(* IEC 61131-3 sources: plc-vscode/tests/st/test-ready/trust-platform/examples/OSCAT/tank_level_pid/non-oop/src, 3 files *)

(* ---- Configuration.st ---- *)
CONFIGURATION TankLevelPidClassicConfiguration
RESOURCE Cpu0 ON PLC
    TASK MainTask (INTERVAL := T#100ms, PRIORITY := 1);
    PROGRAM Main WITH MainTask : Main;
END_RESOURCE
END_CONFIGURATION

(* ---- Main.st ---- *)
PROGRAM Main
VAR
    TankController : CTRL_PID;
    LevelPercent : REAL := REAL#42.0;
    TargetLevelPercent : REAL := REAL#75.0;
    ValveCommandPercent : REAL;
    CommandLimited : BOOL;
END_VAR

TankController(
    ACT := LevelPercent,
    SET_POINT := TargetLevelPercent,
    SUP := REAL#0.0,
    OFS := REAL#0.0,
    M_I := REAL#35.0,
    MAN := TRUE,
    RST := FALSE,
    KP := REAL#2.0,
    TN := REAL#1.0,
    TV := REAL#0.0,
    LL := REAL#0.0,
    LH := REAL#100.0
);
ValveCommandPercent := TankController.Y;
CommandLimited := TankController.LIM;
END_PROGRAM

(* ---- Tests.st ---- *)
TEST_PROGRAM TankLevelPidClassicUsesOscatPidDirectly
VAR
    TankController : CTRL_PID;
END_VAR

TankController(
    ACT := REAL#42.0,
    SET_POINT := REAL#75.0,
    SUP := REAL#0.0,
    OFS := REAL#0.0,
    M_I := REAL#35.0,
    MAN := TRUE,
    RST := FALSE,
    KP := REAL#2.0,
    TN := REAL#1.0,
    TV := REAL#0.0,
    LL := REAL#0.0,
    LH := REAL#100.0
);

ASSERT_NEAR(EXPECTED := REAL#35.0, ACTUAL := TankController.Y, DELTA := REAL#0.001);
ASSERT_FALSE(IN := TankController.LIM);
END_TEST_PROGRAM
